(* IEC 61131-3 sources: Gen-AI/final/Gen-AI_v1.0_submission/A2_框架源码/agent/logs/full34_fixture/E3_P12_1_42/tools/candidate_1/fixture_compile, 1 file *)

(* ---- source.st ---- *)
FUNCTION_BLOCK FB_P12
VAR_INPUT
    THICKNESS_FAULT : BOOL;
    THICKNESS_SIGNAL_VALID : BOOL;
    CUTTING_RUN : BOOL;
    FaultTimestamp : DINT;
    CycleTime : TIME;
END_VAR
VAR_OUTPUT
    THICKNESS_ALARM : BOOL;
    Slab_Fault_Counter : UINT;
    Slab_Runtime_Accumulator : LTIME;
    Slab_Fault_History : ARRAY[0..4] OF DINT;
END_VAR
(* Add a VAR block for internal state/timers before the implementation, if needed. *)
(* SKELETON ONLY: replace this RETURN with scan logic and required initial state. *)
RETURN;
END_FUNCTION_BLOCK

(* FIXTURE_COMPILE_FAIL *)
